% RSLogix 500 project PROGRAM 10.RSS, saved by version 8.30.00.16 %
PROJECT "UNTITLED"    % processor: Bul.1763 MicroLogix 1100 Series B %

PROGRAM FILES
  LAD 2 "MAIN"  4 rungs
  LAD 3 "IO"  10 rungs
  LAD 4 "CONTROLS"  9 rungs
  LAD 5 "ALARMS"  8 rungs

DATA FILES
  O0 OUTPUT  4 elements
  I1 INPUT  6 elements
  S2 STATUS  66 elements
  B3 BINARY  2 elements
  T4 TIMER  4 elements
  C5 COUNTER  1 elements
  R6 CONTROL  1 elements
  N7 INTEGER  3 elements
  F8 FLOAT  1 elements

LADDER 2 "MAIN"
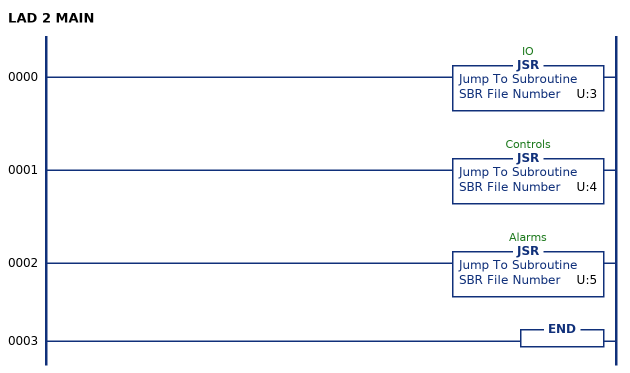
% Rung: 0 %
SOR JSR U:3 EOR
%   U:3  "IO" %
% Rung: 1 %
SOR JSR U:4 EOR
%   U:4  "Controls" %
% Rung: 2 %
SOR JSR U:5 EOR
%   U:5  "Alarms" %
% Rung: 3 %
SOR END EOR

LADDER 3 "IO"
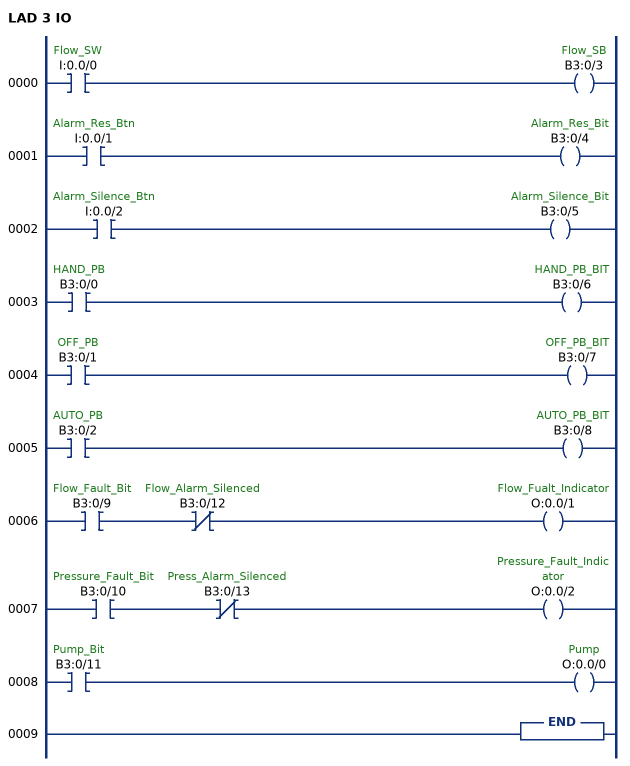
% Rung: 0 %
SOR XIC I:0.0/0 OTE B3:0/3 EOR
%   I:0.0/0  "Flow_SW" %
%   B3:0/3  "Flow_SB" %
% Rung: 1 %
SOR XIC I:0.0/1 OTE B3:0/4 EOR
%   I:0.0/1  "Alarm_Res_Btn" %
%   B3:0/4  "Alarm_Res_Bit" %
% Rung: 2 %
SOR XIC I:0.0/2 OTE B3:0/5 EOR
%   I:0.0/2  "Alarm_Silence_Btn" %
%   B3:0/5  "Alarm_Silence_Bit" %
% Rung: 3 %
SOR XIC B3:0/0 OTE B3:0/6 EOR
%   B3:0/0  "HAND_PB" %
%   B3:0/6  "HAND_PB_BIT" %
% Rung: 4 %
SOR XIC B3:0/1 OTE B3:0/7 EOR
%   B3:0/1  "OFF_PB" %
%   B3:0/7  "OFF_PB_BIT" %
% Rung: 5 %
SOR XIC B3:0/2 OTE B3:0/8 EOR
%   B3:0/2  "AUTO_PB" %
%   B3:0/8  "AUTO_PB_BIT" %
% Rung: 6 %
SOR XIC B3:0/9 XIO B3:0/12 OTE O:0.0/1 EOR
%   B3:0/9  "Flow_Fault_Bit" %
%   B3:0/12  "Flow_Alarm_Silenced" %
%   O:0.0/1  "Flow_Fualt_Indicator" %
% Rung: 7 %
SOR XIC B3:0/10 XIO B3:0/13 OTE O:0.0/2 EOR
%   B3:0/10  "Pressure_Fault_Bit" %
%   B3:0/13  "Press_Alarm_Silenced" %
%   O:0.0/2  "Pressure_Fault_Indic ator" %
% Rung: 8 %
SOR XIC B3:0/11 OTE O:0.0/0 EOR
%   B3:0/11  "Pump_Bit" %
%   O:0.0/0  "Pump" %
% Rung: 9 %
SOR END EOR

LADDER 4 "CONTROLS"
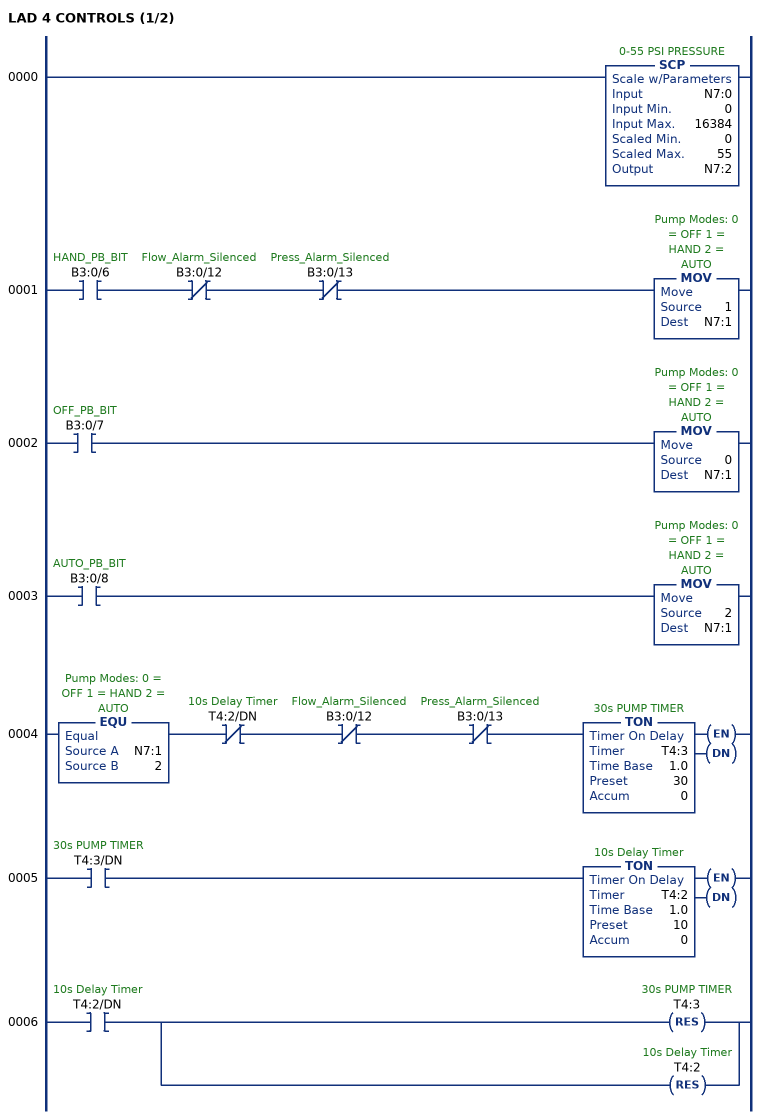
% Rung: 0 %
SOR SCP N7:0 0 16384 0 55 N7:2 EOR
%   N7:0  "Pressure_Sensor" %
%   N7:2  "0-55 PSI PRESSURE" %
% Rung: 1 %
SOR XIC B3:0/6 XIO B3:0/12 XIO B3:0/13 MOV 1 N7:1 EOR
%   B3:0/6  "HAND_PB_BIT" %
%   B3:0/12  "Flow_Alarm_Silenced" %
%   B3:0/13  "Press_Alarm_Silenced" %
%   N7:1  "Pump Modes: 0 = OFF 1 = HAND 2 = AUTO" %
% Rung: 2 %
SOR XIC B3:0/7 MOV 0 N7:1 EOR
%   B3:0/7  "OFF_PB_BIT" %
%   N7:1  "Pump Modes: 0 = OFF 1 = HAND 2 = AUTO" %
% Rung: 3 %
SOR XIC B3:0/8 MOV 2 N7:1 EOR
%   B3:0/8  "AUTO_PB_BIT" %
%   N7:1  "Pump Modes: 0 = OFF 1 = HAND 2 = AUTO" %
% Rung: 4 %
SOR EQU N7:1 2 XIO T4:2/DN XIO B3:0/12 XIO B3:0/13 TON T4:3 1.0 30 0 EOR
%   N7:1  "Pump Modes: 0 = OFF 1 = HAND 2 = AUTO" %
%   T4:2  "10s Delay Timer" %
%   B3:0/12  "Flow_Alarm_Silenced" %
%   B3:0/13  "Press_Alarm_Silenced" %
%   T4:3  "30s PUMP TIMER" %
% Rung: 5 %
SOR XIC T4:3/DN TON T4:2 1.0 10 0 EOR
%   T4:3  "30s PUMP TIMER" %
%   T4:2  "10s Delay Timer" %
% Rung: 6 %
SOR XIC T4:2/DN BST RES T4:3 NXB RES T4:2 BND EOR
%   T4:2  "10s Delay Timer" %
%   T4:3  "30s PUMP TIMER" %

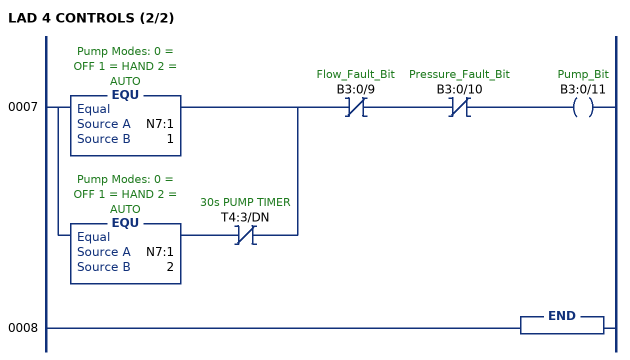
% Rung: 7 %
SOR BST EQU N7:1 1 NXB EQU N7:1 2 XIO T4:3/DN BND XIO B3:0/9 XIO B3:0/10 OTE B3:0/11 EOR
%   N7:1  "Pump Modes: 0 = OFF 1 = HAND 2 = AUTO" %
%   T4:3  "30s PUMP TIMER" %
%   B3:0/9  "Flow_Fault_Bit" %
%   B3:0/10  "Pressure_Fault_Bit" %
%   B3:0/11  "Pump_Bit" %
% Rung: 8 %
SOR END EOR

LADDER 5 "ALARMS"
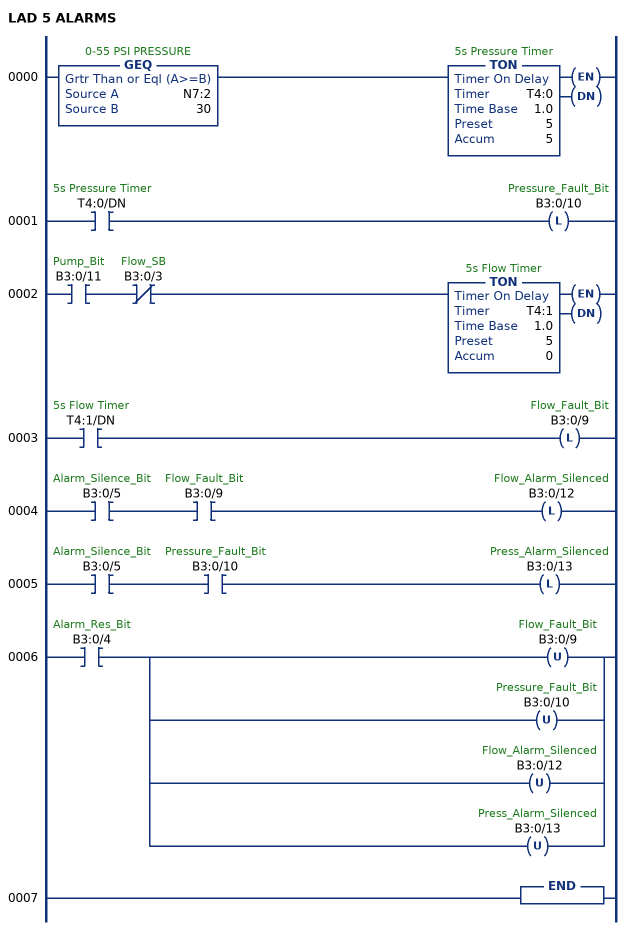
% Rung: 0 %
SOR GEQ N7:2 30 TON T4:0 1.0 5 5 EOR
%   N7:2  "0-55 PSI PRESSURE" %
%   T4:0  "5s Pressure Timer" %
% Rung: 1 %
SOR XIC T4:0/DN OTL B3:0/10 EOR
%   T4:0  "5s Pressure Timer" %
%   B3:0/10  "Pressure_Fault_Bit" %
% Rung: 2 %
SOR XIC B3:0/11 XIO B3:0/3 TON T4:1 1.0 5 0 EOR
%   B3:0/11  "Pump_Bit" %
%   B3:0/3  "Flow_SB" %
%   T4:1  "5s Flow Timer" %
% Rung: 3 %
SOR XIC T4:1/DN OTL B3:0/9 EOR
%   T4:1  "5s Flow Timer" %
%   B3:0/9  "Flow_Fault_Bit" %
% Rung: 4 %
SOR XIC B3:0/5 XIC B3:0/9 OTL B3:0/12 EOR
%   B3:0/5  "Alarm_Silence_Bit" %
%   B3:0/9  "Flow_Fault_Bit" %
%   B3:0/12  "Flow_Alarm_Silenced" %
% Rung: 5 %
SOR XIC B3:0/5 XIC B3:0/10 OTL B3:0/13 EOR
%   B3:0/5  "Alarm_Silence_Bit" %
%   B3:0/10  "Pressure_Fault_Bit" %
%   B3:0/13  "Press_Alarm_Silenced" %
% Rung: 6 %
SOR XIC B3:0/4 BST OTU B3:0/9 NXB OTU B3:0/10 NXB OTU B3:0/12 NXB OTU B3:0/13 BND EOR
%   B3:0/4  "Alarm_Res_Bit" %
%   B3:0/9  "Flow_Fault_Bit" %
%   B3:0/10  "Pressure_Fault_Bit" %
%   B3:0/12  "Flow_Alarm_Silenced" %
%   B3:0/13  "Press_Alarm_Silenced" %
% Rung: 7 %
SOR END EOR

OTHER DOCUMENTED ADDRESSES
  B1:0/0  "Trigger_Alarm_Bit"
  B1:0/2  "ONS"
  B1:0/3  "Alarm_Bit"
  B1:0/4  "ONS"
  B3:0/14  "ONS"
  B3:1/3  "ONS"

DATA TABLE (non-zero values as saved)
DATA B3
% B3:0 % 0X4048 0X0000
DATA T4
% .PRE .ACC %
% T4:0 % 5 5
% T4:1 % 5 0
% T4:2 % 10 0
% T4:3 % 30 0
DATA N7
% N7:0 % 10000 1 34
